// TIA Portal V20 export
DATA_BLOCK "DB_HMI_recype"   // DB2
{ S7_Optimized_Access := 'TRUE' }
// stored: MemoryReserve 100
   VAR
      recipe : Struct
         Zprava : Int := 2;   // dvoumístné číslo přeneseno a doplněno po bytech do šablony zprávy
         PRG_CAM_etiketa : Int := 1;   // program v kameře která kontroluje papír co se vkládá pod folii
         PRG_CAM_folie : Int;   // kamery kontrolující folii
         vyrazovac_on_off : Bool := true;   // false - neposílat signál pro vyřazovač
         variabilni_pole_on_off : Bool := true;   // false - neposílat variabilní pole
         pole_string_1 : String[20] := 'Ceska republika';   // textove_pole - není bráno z receptůry ale volně zadatalné
         pole_string_2 : String[10];   // textove_pole - není bráno z receptůry ale volně zadatalné
      END_STRUCT;
      fronta : Array[1..5] of Struct
         prenaseny_text : String[100];   // načtený text kamerou
         balik_den : Int;   // aktualni číslo plata
         vyrazeni : Bool;   // vyřazení
      END_STRUCT;
      obsazenost_fronty : Int;
      ODESLI_dATA : Bool;
      VZDALENOST_KAMERA_ETIKETA_POZADOVANA : DInt := 20;
      VZDALENOST_KAMERY_FOLIE_POZADOVANA : DInt := 150;
      meze : DInt := 35;
      aktualni_poloha : DInt;
   END_VAR
BEGIN
END_DATA_BLOCK
